(* IEC 61131-3 sources: codesys-build/examples/frame-assembly/src/generated/types/ST_LineCS1001, 3 files *)

(* ---- ST_LineCS1001.st ---- *)
(*
Auxiliary control signals and feedback for an Intelligrated CS1001 motor-driven roller card.
https://www.scribd.com/document/823553754/MDR-710-With-WWL-Installation-and-Maintenance-Manual
*)
TYPE ST_LineCS1001 :
STRUCT
	(* Normalized auxiliary control signals toward one card; mapping handles electrical polarity. *)
	Output : ST_LineCS1001Output;
	(* Digital feedback from the CS1001 auxiliary terminals, interpreted using the configured signal polarity. *)
	Input : ST_LineCS1001Input;
END_STRUCT
END_TYPE

(* ---- ST_LineCS1001Input.st ---- *)
(*
Auxiliary control signals and feedback for an Intelligrated CS1001 motor-driven roller card.
https://www.scribd.com/document/823553754/MDR-710-With-WWL-Installation-and-Maintenance-Manual
*)
TYPE ST_LineCS1001Input :
STRUCT
	(* CN2-4 sensor indication; TRUE when the photoeye is blocked. *)
	Sensor : BOOL;
	(* CN2-5 aggregate error indication; no numeric diagnostic code is transmitted by this bit. *)
	Error : BOOL;
	(* CN2-6 warning indication. *)
	Warning : BOOL;
	(* CN2-7 synchronization indication; TRUE indicates motor running after polarity conversion. *)
	Sync : BOOL;
END_STRUCT
END_TYPE

(* ---- ST_LineCS1001Output.st ---- *)
(*
Auxiliary control signals and feedback for an Intelligrated CS1001 motor-driven roller card.
https://www.scribd.com/document/823553754/MDR-710-With-WWL-Installation-and-Maintenance-Manual
*)
TYPE ST_LineCS1001Output :
STRUCT
	(* Assert CN2-1 according to the installed SW2-6 setting. TRUE can force run or hold accumulation; FALSE can release accumulation. *)
	MotionAsserted : BOOL;
	(* CN2-2 role depends on card mode. Do not interpret as left/right diverter routing. *)
	DirectionOrSlaveErrorAsserted : BOOL;
	(* Optional CN2-3 reference in 0..10 V. Not metres/second and not a 4..20 mA signal. *)
	SpeedVolts : LREAL;
END_STRUCT
END_TYPE
